Fanuc KAREL source: KO00031.KL

PROGRAM KO00031
%NOLOCKGROUP
VAR
  P1: JOINTPOS
  P2: JOINTPOS
  P3: JOINTPOS
  P4: JOINTPOS
  OUT: XYZWPREXT
BEGIN
  OUT = FRAME(P1, P2, P3, P4)
END KO00031
